TYPE ST_Piston_SelectionList :
STRUCT
	Num: INT;
	Description: STRING(80);

END_STRUCT
END_TYPE

(* stored: Version 1.1.0.1, ProductVersion 3.1.4024.12
   DUT ST_Piston_SelectionList: Id {4b2d3383-913f-41f7-8325-d999225275db} *)
